(* IEC 61131-3 sources: SemantiST/compiler/intake/normalize/probes/scl-organization-block, 2 files *)

(* ---- original.st ---- *)
ORGANIZATION_BLOCK CYCLE
VAR
    N : INT;
END_VAR
N := N + 1;
END_ORGANIZATION_BLOCK

FUNCTION main : DINT
CYCLE(); CYCLE();
printf('%d$N', CYCLE.N);
main := 0;
END_FUNCTION

(* ---- rewritten.st ---- *)
PROGRAM CYCLE
VAR
    N : INT;
END_VAR
N := N + 1;
END_PROGRAM

FUNCTION main : DINT
CYCLE(); CYCLE();
printf('%d$N', CYCLE.N);
main := 0;
END_FUNCTION
